Fanuc KAREL source: kt00896.KL

-- PROVISIONAL review KL for V1013-1; original PC SHA256 0fcac0dd3cd1cadf09860e91820669934179603e577e1b5a633d0430b73fca11
-- Incomplete behavior may be omitted. Consult companion uncertainty JSON. Do not deploy.
PROGRAM KT00896
%NOLOCKGROUP
VAR
  OUT : BOOLEAN
-- UNRESOLVED_DECL P1 type=000199
-- UNRESOLVED_DECL P2 type=000199
BEGIN
  -- UNRESOLVED_PC offsets 5-31; opcodes 27,27,49,7E,AD,27,9D,76,23
  -- UNRESOLVED_PC offsets 36-40; opcodes 7F
END KT00896
